TYPE ST_HW_DO :
STRUCT
END_STRUCT
END_TYPE

(* stored: Version 1.1.0.1, ProductVersion 3.1.4024.13
   DUT ST_HW_DO: Id {35f9c9cd-d985-4075-9b90-95c672f87b3b} *)
